{attribute 'qualified_only'}
VAR_GLOBAL
	parameters	: TYPE_PARAMETERS;
	homing		: TYPE_SEQUENCE;
	sequence	: ARRAY[0..Size.MAX_SEQUENCE-1] OF TYPE_SEQUENCE;
	prgState	: PRGSTATE_ENUM;
END_VAR

(* stored: Version 1.1.0.1, ProductVersion 3.1.4024.12
   GVL ProgramDB: Id {fcf68a51-2b91-462e-8ddc-f45260ef6fb1} *)
